# EPICS substitutions: db/Beckhoff_7XXX/ecmcEP7211-0034_OPT_csv.substitutions
file "ecmcEL72XX_DRV.template"
{
  pattern {CH_ID}
          {01   }
}
